{attribute 'qualified_only'}
VAR_GLOBAL CONSTANT
    cMaxLights : UINT := 16;
    cMaxButtons : UINT := 16;
END_VAR

(* stored: Version 1.1.0.1
   GVL GVL_HomeLimits: Id {c7dd2490-1ccc-4b72-a1a2-a20db484e5db} *)
